// TIA Portal V19 export
FUNCTION "PID_DATA_MAPPING" : Void   // FC3, LAD
{ S7_Optimized_Access := 'TRUE' }
// stored: SetENOAutomatically false
BEGIN

REGION Network 1: -------------------------------------------------- REACTOR-1 ------------------------------------------------------------------
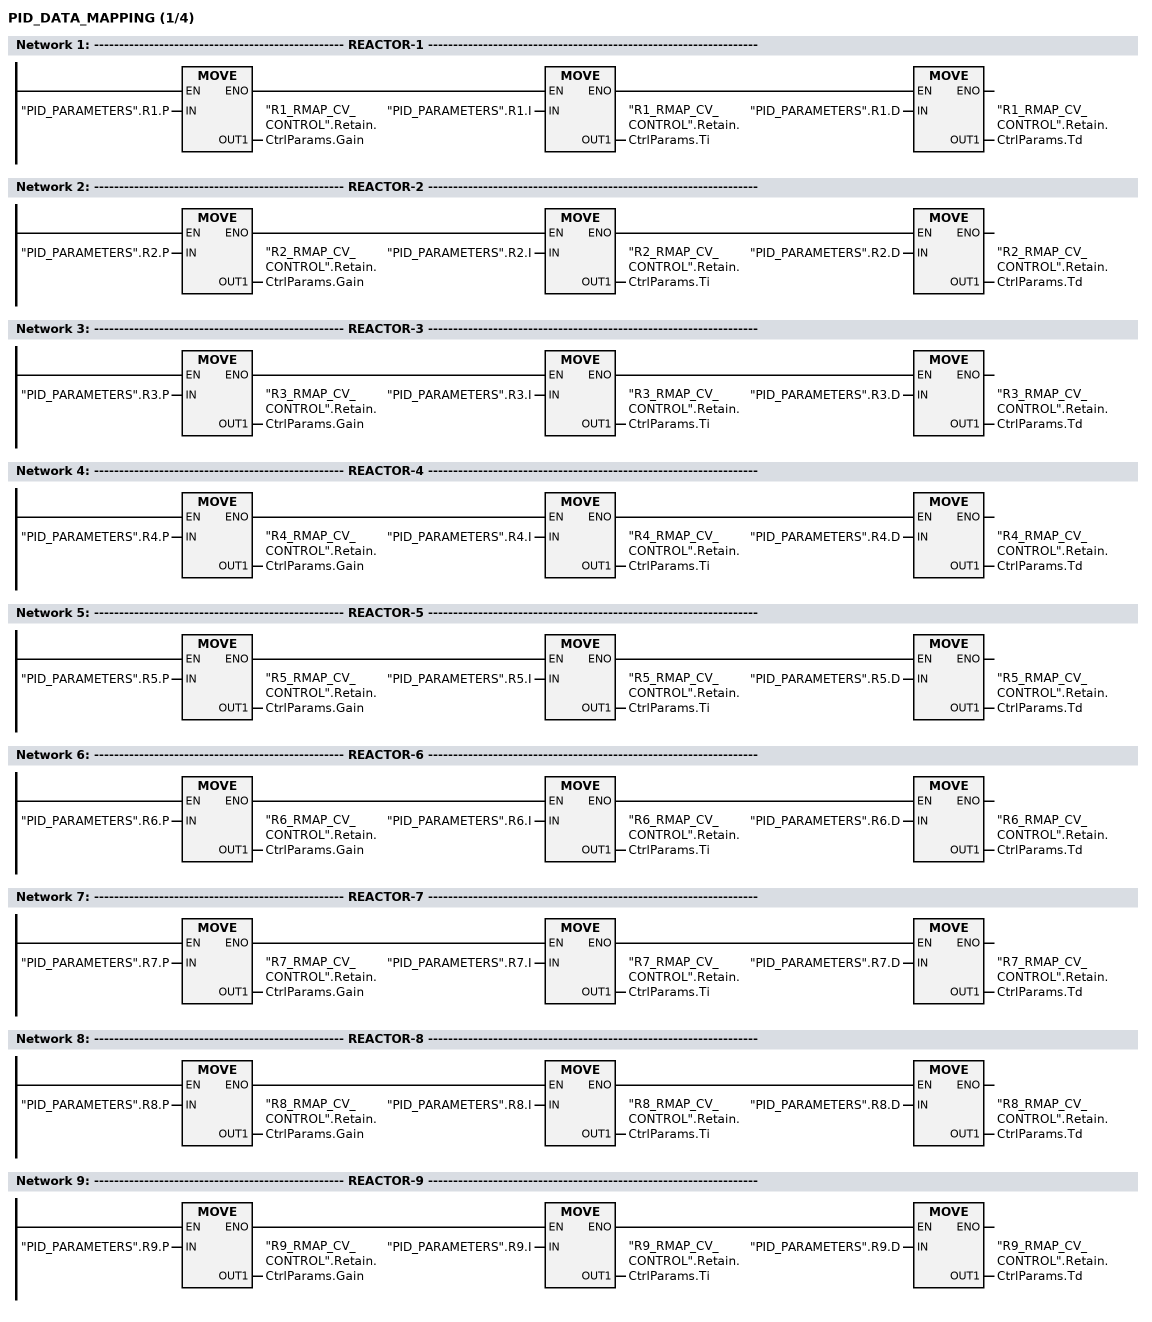
   RUNG wire#powerrail
      Move(in := "PID_PARAMETERS".R1.P, out1 => "R1_RMAP_CV_CONTROL".Retain.CtrlParams.Gain)
      Move(in := "PID_PARAMETERS".R1.I, out1 => "R1_RMAP_CV_CONTROL".Retain.CtrlParams.Ti)
      Move(in := "PID_PARAMETERS".R1.D, out1 => "R1_RMAP_CV_CONTROL".Retain.CtrlParams.Td)
   END_RUNG
   // the same network as SCL:
   "R1_RMAP_CV_CONTROL".Retain.CtrlParams.Gain := "PID_PARAMETERS".R1.P;
   "R1_RMAP_CV_CONTROL".Retain.CtrlParams.Ti := "PID_PARAMETERS".R1.I;
   "R1_RMAP_CV_CONTROL".Retain.CtrlParams.Td := "PID_PARAMETERS".R1.D;
END_REGION

REGION Network 2: -------------------------------------------------- REACTOR-2 ------------------------------------------------------------------
   RUNG wire#powerrail
      Move(in := "PID_PARAMETERS".R2.P, out1 => "R2_RMAP_CV_CONTROL".Retain.CtrlParams.Gain)
      Move(in := "PID_PARAMETERS".R2.I, out1 => "R2_RMAP_CV_CONTROL".Retain.CtrlParams.Ti)
      Move(in := "PID_PARAMETERS".R2.D, out1 => "R2_RMAP_CV_CONTROL".Retain.CtrlParams.Td)
   END_RUNG
   // the same network as SCL:
   "R2_RMAP_CV_CONTROL".Retain.CtrlParams.Gain := "PID_PARAMETERS".R2.P;
   "R2_RMAP_CV_CONTROL".Retain.CtrlParams.Ti := "PID_PARAMETERS".R2.I;
   "R2_RMAP_CV_CONTROL".Retain.CtrlParams.Td := "PID_PARAMETERS".R2.D;
END_REGION

REGION Network 3: -------------------------------------------------- REACTOR-3 ------------------------------------------------------------------
   RUNG wire#powerrail
      Move(in := "PID_PARAMETERS".R3.P, out1 => "R3_RMAP_CV_CONTROL".Retain.CtrlParams.Gain)
      Move(in := "PID_PARAMETERS".R3.I, out1 => "R3_RMAP_CV_CONTROL".Retain.CtrlParams.Ti)
      Move(in := "PID_PARAMETERS".R3.D, out1 => "R3_RMAP_CV_CONTROL".Retain.CtrlParams.Td)
   END_RUNG
   // the same network as SCL:
   "R3_RMAP_CV_CONTROL".Retain.CtrlParams.Gain := "PID_PARAMETERS".R3.P;
   "R3_RMAP_CV_CONTROL".Retain.CtrlParams.Ti := "PID_PARAMETERS".R3.I;
   "R3_RMAP_CV_CONTROL".Retain.CtrlParams.Td := "PID_PARAMETERS".R3.D;
END_REGION

REGION Network 4: -------------------------------------------------- REACTOR-4 ------------------------------------------------------------------
   RUNG wire#powerrail
      Move(in := "PID_PARAMETERS".R4.P, out1 => "R4_RMAP_CV_CONTROL".Retain.CtrlParams.Gain)
      Move(in := "PID_PARAMETERS".R4.I, out1 => "R4_RMAP_CV_CONTROL".Retain.CtrlParams.Ti)
      Move(in := "PID_PARAMETERS".R4.D, out1 => "R4_RMAP_CV_CONTROL".Retain.CtrlParams.Td)
   END_RUNG
   // the same network as SCL:
   "R4_RMAP_CV_CONTROL".Retain.CtrlParams.Gain := "PID_PARAMETERS".R4.P;
   "R4_RMAP_CV_CONTROL".Retain.CtrlParams.Ti := "PID_PARAMETERS".R4.I;
   "R4_RMAP_CV_CONTROL".Retain.CtrlParams.Td := "PID_PARAMETERS".R4.D;
END_REGION

REGION Network 5: -------------------------------------------------- REACTOR-5 ------------------------------------------------------------------
   RUNG wire#powerrail
      Move(in := "PID_PARAMETERS".R5.P, out1 => "R5_RMAP_CV_CONTROL".Retain.CtrlParams.Gain)
      Move(in := "PID_PARAMETERS".R5.I, out1 => "R5_RMAP_CV_CONTROL".Retain.CtrlParams.Ti)
      Move(in := "PID_PARAMETERS".R5.D, out1 => "R5_RMAP_CV_CONTROL".Retain.CtrlParams.Td)
   END_RUNG
   // the same network as SCL:
   "R5_RMAP_CV_CONTROL".Retain.CtrlParams.Gain := "PID_PARAMETERS".R5.P;
   "R5_RMAP_CV_CONTROL".Retain.CtrlParams.Ti := "PID_PARAMETERS".R5.I;
   "R5_RMAP_CV_CONTROL".Retain.CtrlParams.Td := "PID_PARAMETERS".R5.D;
END_REGION

REGION Network 6: -------------------------------------------------- REACTOR-6 ------------------------------------------------------------------
   RUNG wire#powerrail
      Move(in := "PID_PARAMETERS".R6.P, out1 => "R6_RMAP_CV_CONTROL".Retain.CtrlParams.Gain)
      Move(in := "PID_PARAMETERS".R6.I, out1 => "R6_RMAP_CV_CONTROL".Retain.CtrlParams.Ti)
      Move(in := "PID_PARAMETERS".R6.D, out1 => "R6_RMAP_CV_CONTROL".Retain.CtrlParams.Td)
   END_RUNG
   // the same network as SCL:
   "R6_RMAP_CV_CONTROL".Retain.CtrlParams.Gain := "PID_PARAMETERS".R6.P;
   "R6_RMAP_CV_CONTROL".Retain.CtrlParams.Ti := "PID_PARAMETERS".R6.I;
   "R6_RMAP_CV_CONTROL".Retain.CtrlParams.Td := "PID_PARAMETERS".R6.D;
END_REGION

REGION Network 7: -------------------------------------------------- REACTOR-7 ------------------------------------------------------------------
   RUNG wire#powerrail
      Move(in := "PID_PARAMETERS".R7.P, out1 => "R7_RMAP_CV_CONTROL".Retain.CtrlParams.Gain)
      Move(in := "PID_PARAMETERS".R7.I, out1 => "R7_RMAP_CV_CONTROL".Retain.CtrlParams.Ti)
      Move(in := "PID_PARAMETERS".R7.D, out1 => "R7_RMAP_CV_CONTROL".Retain.CtrlParams.Td)
   END_RUNG
   // the same network as SCL:
   "R7_RMAP_CV_CONTROL".Retain.CtrlParams.Gain := "PID_PARAMETERS".R7.P;
   "R7_RMAP_CV_CONTROL".Retain.CtrlParams.Ti := "PID_PARAMETERS".R7.I;
   "R7_RMAP_CV_CONTROL".Retain.CtrlParams.Td := "PID_PARAMETERS".R7.D;
END_REGION

REGION Network 8: -------------------------------------------------- REACTOR-8 ------------------------------------------------------------------
   RUNG wire#powerrail
      Move(in := "PID_PARAMETERS".R8.P, out1 => "R8_RMAP_CV_CONTROL".Retain.CtrlParams.Gain)
      Move(in := "PID_PARAMETERS".R8.I, out1 => "R8_RMAP_CV_CONTROL".Retain.CtrlParams.Ti)
      Move(in := "PID_PARAMETERS".R8.D, out1 => "R8_RMAP_CV_CONTROL".Retain.CtrlParams.Td)
   END_RUNG
   // the same network as SCL:
   "R8_RMAP_CV_CONTROL".Retain.CtrlParams.Gain := "PID_PARAMETERS".R8.P;
   "R8_RMAP_CV_CONTROL".Retain.CtrlParams.Ti := "PID_PARAMETERS".R8.I;
   "R8_RMAP_CV_CONTROL".Retain.CtrlParams.Td := "PID_PARAMETERS".R8.D;
END_REGION

REGION Network 9: -------------------------------------------------- REACTOR-9 ------------------------------------------------------------------
   RUNG wire#powerrail
      Move(in := "PID_PARAMETERS".R9.P, out1 => "R9_RMAP_CV_CONTROL".Retain.CtrlParams.Gain)
      Move(in := "PID_PARAMETERS".R9.I, out1 => "R9_RMAP_CV_CONTROL".Retain.CtrlParams.Ti)
      Move(in := "PID_PARAMETERS".R9.D, out1 => "R9_RMAP_CV_CONTROL".Retain.CtrlParams.Td)
   END_RUNG
   // the same network as SCL:
   "R9_RMAP_CV_CONTROL".Retain.CtrlParams.Gain := "PID_PARAMETERS".R9.P;
   "R9_RMAP_CV_CONTROL".Retain.CtrlParams.Ti := "PID_PARAMETERS".R9.I;
   "R9_RMAP_CV_CONTROL".Retain.CtrlParams.Td := "PID_PARAMETERS".R9.D;
END_REGION

REGION Network 10: -------------------------------------------------- REACTOR-10 ------------------------------------------------------------------
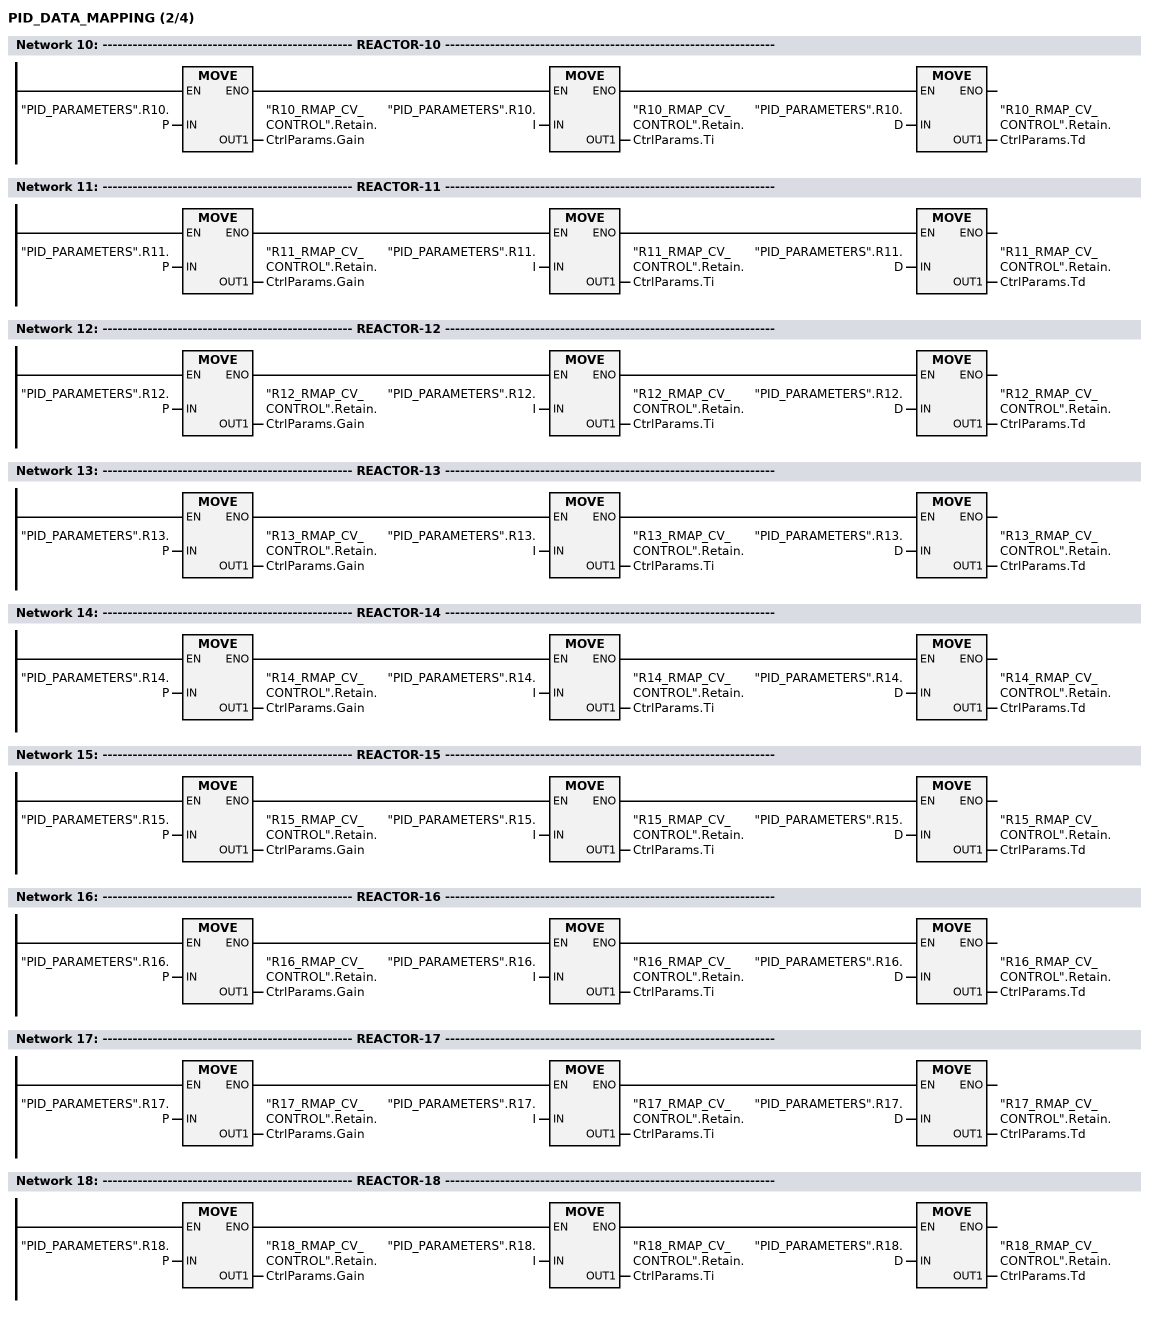
   RUNG wire#powerrail
      Move(in := "PID_PARAMETERS".R10.P, out1 => "R10_RMAP_CV_CONTROL".Retain.CtrlParams.Gain)
      Move(in := "PID_PARAMETERS".R10.I, out1 => "R10_RMAP_CV_CONTROL".Retain.CtrlParams.Ti)
      Move(in := "PID_PARAMETERS".R10.D, out1 => "R10_RMAP_CV_CONTROL".Retain.CtrlParams.Td)
   END_RUNG
   // the same network as SCL:
   "R10_RMAP_CV_CONTROL".Retain.CtrlParams.Gain := "PID_PARAMETERS".R10.P;
   "R10_RMAP_CV_CONTROL".Retain.CtrlParams.Ti := "PID_PARAMETERS".R10.I;
   "R10_RMAP_CV_CONTROL".Retain.CtrlParams.Td := "PID_PARAMETERS".R10.D;
END_REGION

REGION Network 11: -------------------------------------------------- REACTOR-11 ------------------------------------------------------------------
   RUNG wire#powerrail
      Move(in := "PID_PARAMETERS".R11.P, out1 => "R11_RMAP_CV_CONTROL".Retain.CtrlParams.Gain)
      Move(in := "PID_PARAMETERS".R11.I, out1 => "R11_RMAP_CV_CONTROL".Retain.CtrlParams.Ti)
      Move(in := "PID_PARAMETERS".R11.D, out1 => "R11_RMAP_CV_CONTROL".Retain.CtrlParams.Td)
   END_RUNG
   // the same network as SCL:
   "R11_RMAP_CV_CONTROL".Retain.CtrlParams.Gain := "PID_PARAMETERS".R11.P;
   "R11_RMAP_CV_CONTROL".Retain.CtrlParams.Ti := "PID_PARAMETERS".R11.I;
   "R11_RMAP_CV_CONTROL".Retain.CtrlParams.Td := "PID_PARAMETERS".R11.D;
END_REGION

REGION Network 12: -------------------------------------------------- REACTOR-12 ------------------------------------------------------------------
   RUNG wire#powerrail
      Move(in := "PID_PARAMETERS".R12.P, out1 => "R12_RMAP_CV_CONTROL".Retain.CtrlParams.Gain)
      Move(in := "PID_PARAMETERS".R12.I, out1 => "R12_RMAP_CV_CONTROL".Retain.CtrlParams.Ti)
      Move(in := "PID_PARAMETERS".R12.D, out1 => "R12_RMAP_CV_CONTROL".Retain.CtrlParams.Td)
   END_RUNG
   // the same network as SCL:
   "R12_RMAP_CV_CONTROL".Retain.CtrlParams.Gain := "PID_PARAMETERS".R12.P;
   "R12_RMAP_CV_CONTROL".Retain.CtrlParams.Ti := "PID_PARAMETERS".R12.I;
   "R12_RMAP_CV_CONTROL".Retain.CtrlParams.Td := "PID_PARAMETERS".R12.D;
END_REGION

REGION Network 13: -------------------------------------------------- REACTOR-13 ------------------------------------------------------------------
   RUNG wire#powerrail
      Move(in := "PID_PARAMETERS".R13.P, out1 => "R13_RMAP_CV_CONTROL".Retain.CtrlParams.Gain)
      Move(in := "PID_PARAMETERS".R13.I, out1 => "R13_RMAP_CV_CONTROL".Retain.CtrlParams.Ti)
      Move(in := "PID_PARAMETERS".R13.D, out1 => "R13_RMAP_CV_CONTROL".Retain.CtrlParams.Td)
   END_RUNG
   // the same network as SCL:
   "R13_RMAP_CV_CONTROL".Retain.CtrlParams.Gain := "PID_PARAMETERS".R13.P;
   "R13_RMAP_CV_CONTROL".Retain.CtrlParams.Ti := "PID_PARAMETERS".R13.I;
   "R13_RMAP_CV_CONTROL".Retain.CtrlParams.Td := "PID_PARAMETERS".R13.D;
END_REGION

REGION Network 14: -------------------------------------------------- REACTOR-14 ------------------------------------------------------------------
   RUNG wire#powerrail
      Move(in := "PID_PARAMETERS".R14.P, out1 => "R14_RMAP_CV_CONTROL".Retain.CtrlParams.Gain)
      Move(in := "PID_PARAMETERS".R14.I, out1 => "R14_RMAP_CV_CONTROL".Retain.CtrlParams.Ti)
      Move(in := "PID_PARAMETERS".R14.D, out1 => "R14_RMAP_CV_CONTROL".Retain.CtrlParams.Td)
   END_RUNG
   // the same network as SCL:
   "R14_RMAP_CV_CONTROL".Retain.CtrlParams.Gain := "PID_PARAMETERS".R14.P;
   "R14_RMAP_CV_CONTROL".Retain.CtrlParams.Ti := "PID_PARAMETERS".R14.I;
   "R14_RMAP_CV_CONTROL".Retain.CtrlParams.Td := "PID_PARAMETERS".R14.D;
END_REGION

REGION Network 15: -------------------------------------------------- REACTOR-15 ------------------------------------------------------------------
   RUNG wire#powerrail
      Move(in := "PID_PARAMETERS".R15.P, out1 => "R15_RMAP_CV_CONTROL".Retain.CtrlParams.Gain)
      Move(in := "PID_PARAMETERS".R15.I, out1 => "R15_RMAP_CV_CONTROL".Retain.CtrlParams.Ti)
      Move(in := "PID_PARAMETERS".R15.D, out1 => "R15_RMAP_CV_CONTROL".Retain.CtrlParams.Td)
   END_RUNG
   // the same network as SCL:
   "R15_RMAP_CV_CONTROL".Retain.CtrlParams.Gain := "PID_PARAMETERS".R15.P;
   "R15_RMAP_CV_CONTROL".Retain.CtrlParams.Ti := "PID_PARAMETERS".R15.I;
   "R15_RMAP_CV_CONTROL".Retain.CtrlParams.Td := "PID_PARAMETERS".R15.D;
END_REGION

REGION Network 16: -------------------------------------------------- REACTOR-16 ------------------------------------------------------------------
   RUNG wire#powerrail
      Move(in := "PID_PARAMETERS".R16.P, out1 => "R16_RMAP_CV_CONTROL".Retain.CtrlParams.Gain)
      Move(in := "PID_PARAMETERS".R16.I, out1 => "R16_RMAP_CV_CONTROL".Retain.CtrlParams.Ti)
      Move(in := "PID_PARAMETERS".R16.D, out1 => "R16_RMAP_CV_CONTROL".Retain.CtrlParams.Td)
   END_RUNG
   // the same network as SCL:
   "R16_RMAP_CV_CONTROL".Retain.CtrlParams.Gain := "PID_PARAMETERS".R16.P;
   "R16_RMAP_CV_CONTROL".Retain.CtrlParams.Ti := "PID_PARAMETERS".R16.I;
   "R16_RMAP_CV_CONTROL".Retain.CtrlParams.Td := "PID_PARAMETERS".R16.D;
END_REGION

REGION Network 17: -------------------------------------------------- REACTOR-17 ------------------------------------------------------------------
   RUNG wire#powerrail
      Move(in := "PID_PARAMETERS".R17.P, out1 => "R17_RMAP_CV_CONTROL".Retain.CtrlParams.Gain)
      Move(in := "PID_PARAMETERS".R17.I, out1 => "R17_RMAP_CV_CONTROL".Retain.CtrlParams.Ti)
      Move(in := "PID_PARAMETERS".R17.D, out1 => "R17_RMAP_CV_CONTROL".Retain.CtrlParams.Td)
   END_RUNG
   // the same network as SCL:
   "R17_RMAP_CV_CONTROL".Retain.CtrlParams.Gain := "PID_PARAMETERS".R17.P;
   "R17_RMAP_CV_CONTROL".Retain.CtrlParams.Ti := "PID_PARAMETERS".R17.I;
   "R17_RMAP_CV_CONTROL".Retain.CtrlParams.Td := "PID_PARAMETERS".R17.D;
END_REGION

REGION Network 18: -------------------------------------------------- REACTOR-18 ------------------------------------------------------------------
   RUNG wire#powerrail
      Move(in := "PID_PARAMETERS".R18.P, out1 => "R18_RMAP_CV_CONTROL".Retain.CtrlParams.Gain)
      Move(in := "PID_PARAMETERS".R18.I, out1 => "R18_RMAP_CV_CONTROL".Retain.CtrlParams.Ti)
      Move(in := "PID_PARAMETERS".R18.D, out1 => "R18_RMAP_CV_CONTROL".Retain.CtrlParams.Td)
   END_RUNG
   // the same network as SCL:
   "R18_RMAP_CV_CONTROL".Retain.CtrlParams.Gain := "PID_PARAMETERS".R18.P;
   "R18_RMAP_CV_CONTROL".Retain.CtrlParams.Ti := "PID_PARAMETERS".R18.I;
   "R18_RMAP_CV_CONTROL".Retain.CtrlParams.Td := "PID_PARAMETERS".R18.D;
END_REGION

REGION Network 19: -------------------------------------------------- HS_CP01 ------------------------------------------------------------------
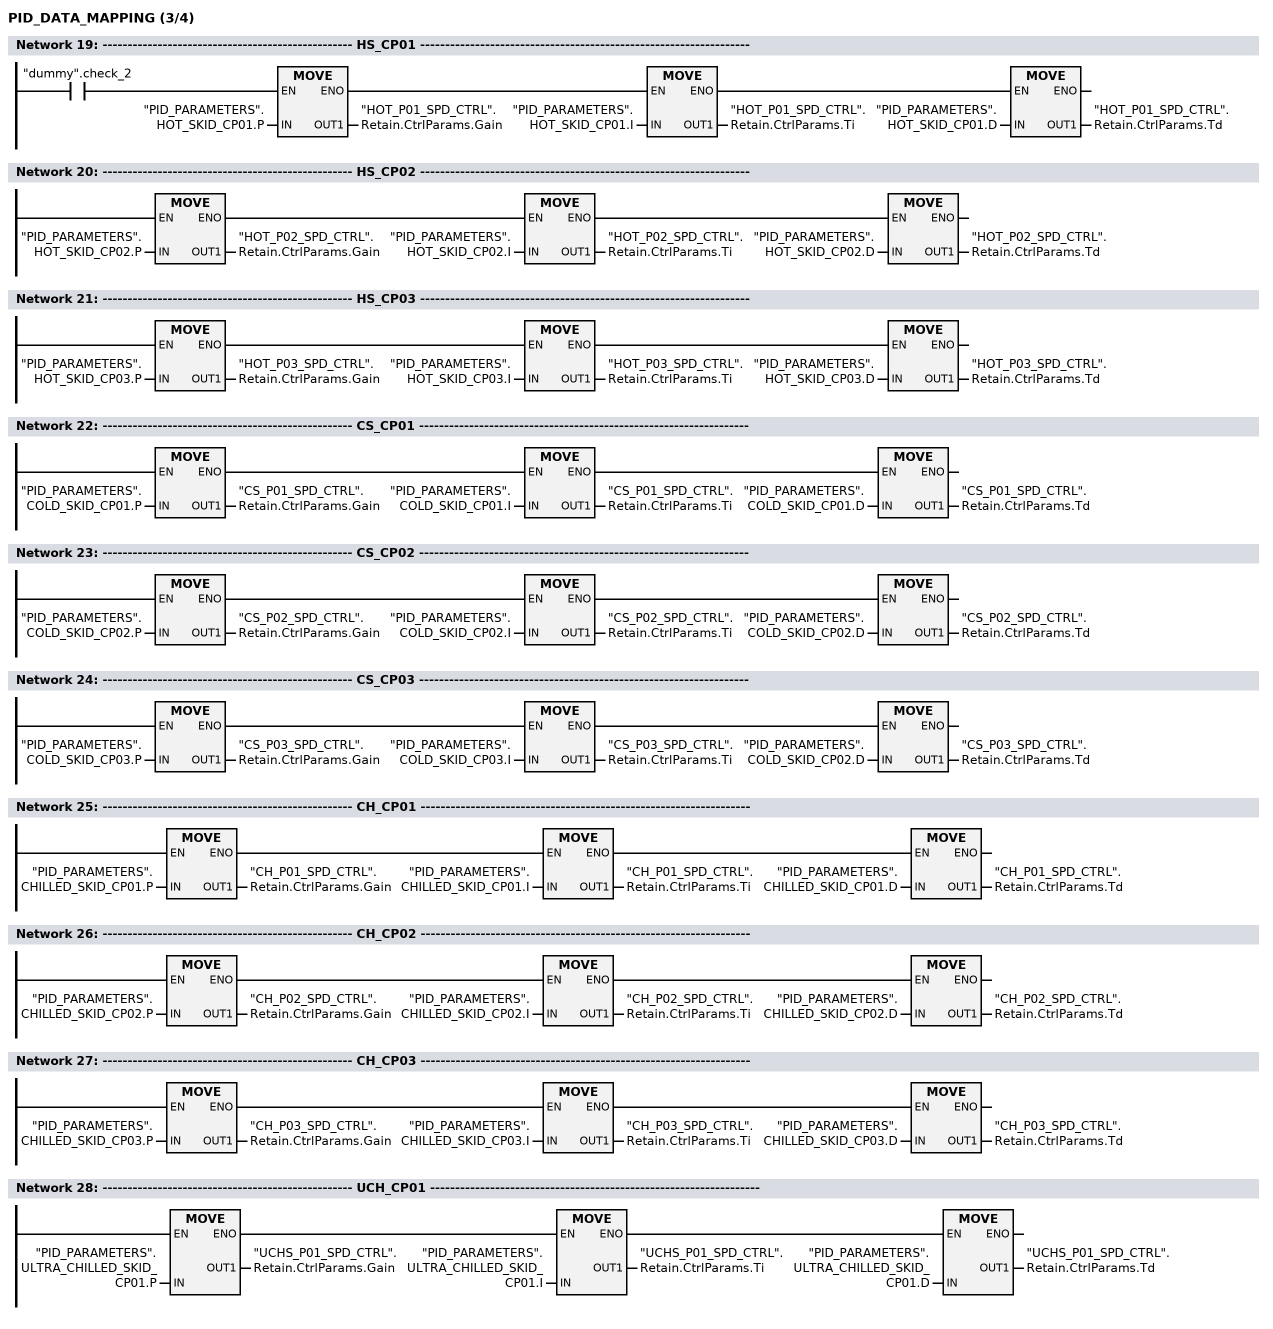
   RUNG wire#powerrail
      Contact( "dummy".check_2 )
      Move(in := "PID_PARAMETERS".HOT_SKID_CP01.P, out1 => "HOT_P01_SPD_CTRL".Retain.CtrlParams.Gain)
      Move(in := "PID_PARAMETERS".HOT_SKID_CP01.I, out1 => "HOT_P01_SPD_CTRL".Retain.CtrlParams.Ti)
      Move(in := "PID_PARAMETERS".HOT_SKID_CP01.D, out1 => "HOT_P01_SPD_CTRL".Retain.CtrlParams.Td)
   END_RUNG
   // the same network as SCL:
   IF "dummy".check_2 THEN
       "HOT_P01_SPD_CTRL".Retain.CtrlParams.Gain := "PID_PARAMETERS".HOT_SKID_CP01.P;
       "HOT_P01_SPD_CTRL".Retain.CtrlParams.Ti := "PID_PARAMETERS".HOT_SKID_CP01.I;
       "HOT_P01_SPD_CTRL".Retain.CtrlParams.Td := "PID_PARAMETERS".HOT_SKID_CP01.D;
   END_IF;
END_REGION

REGION Network 20: -------------------------------------------------- HS_CP02 ------------------------------------------------------------------
   RUNG wire#powerrail
      Move(in := "PID_PARAMETERS".HOT_SKID_CP02.P, out1 => "HOT_P02_SPD_CTRL".Retain.CtrlParams.Gain)
      Move(in := "PID_PARAMETERS".HOT_SKID_CP02.I, out1 => "HOT_P02_SPD_CTRL".Retain.CtrlParams.Ti)
      Move(in := "PID_PARAMETERS".HOT_SKID_CP02.D, out1 => "HOT_P02_SPD_CTRL".Retain.CtrlParams.Td)
   END_RUNG
   // the same network as SCL:
   "HOT_P02_SPD_CTRL".Retain.CtrlParams.Gain := "PID_PARAMETERS".HOT_SKID_CP02.P;
   "HOT_P02_SPD_CTRL".Retain.CtrlParams.Ti := "PID_PARAMETERS".HOT_SKID_CP02.I;
   "HOT_P02_SPD_CTRL".Retain.CtrlParams.Td := "PID_PARAMETERS".HOT_SKID_CP02.D;
END_REGION

REGION Network 21: -------------------------------------------------- HS_CP03 ------------------------------------------------------------------
   RUNG wire#powerrail
      Move(in := "PID_PARAMETERS".HOT_SKID_CP03.P, out1 => "HOT_P03_SPD_CTRL".Retain.CtrlParams.Gain)
      Move(in := "PID_PARAMETERS".HOT_SKID_CP03.I, out1 => "HOT_P03_SPD_CTRL".Retain.CtrlParams.Ti)
      Move(in := "PID_PARAMETERS".HOT_SKID_CP03.D, out1 => "HOT_P03_SPD_CTRL".Retain.CtrlParams.Td)
   END_RUNG
   // the same network as SCL:
   "HOT_P03_SPD_CTRL".Retain.CtrlParams.Gain := "PID_PARAMETERS".HOT_SKID_CP03.P;
   "HOT_P03_SPD_CTRL".Retain.CtrlParams.Ti := "PID_PARAMETERS".HOT_SKID_CP03.I;
   "HOT_P03_SPD_CTRL".Retain.CtrlParams.Td := "PID_PARAMETERS".HOT_SKID_CP03.D;
END_REGION

REGION Network 22: -------------------------------------------------- CS_CP01 ------------------------------------------------------------------
   RUNG wire#powerrail
      Move(in := "PID_PARAMETERS".COLD_SKID_CP01.P, out1 => "CS_P01_SPD_CTRL".Retain.CtrlParams.Gain)
      Move(in := "PID_PARAMETERS".COLD_SKID_CP01.I, out1 => "CS_P01_SPD_CTRL".Retain.CtrlParams.Ti)
      Move(in := "PID_PARAMETERS".COLD_SKID_CP01.D, out1 => "CS_P01_SPD_CTRL".Retain.CtrlParams.Td)
   END_RUNG
   // the same network as SCL:
   "CS_P01_SPD_CTRL".Retain.CtrlParams.Gain := "PID_PARAMETERS".COLD_SKID_CP01.P;
   "CS_P01_SPD_CTRL".Retain.CtrlParams.Ti := "PID_PARAMETERS".COLD_SKID_CP01.I;
   "CS_P01_SPD_CTRL".Retain.CtrlParams.Td := "PID_PARAMETERS".COLD_SKID_CP01.D;
END_REGION

REGION Network 23: -------------------------------------------------- CS_CP02 ------------------------------------------------------------------
   RUNG wire#powerrail
      Move(in := "PID_PARAMETERS".COLD_SKID_CP02.P, out1 => "CS_P02_SPD_CTRL".Retain.CtrlParams.Gain)
      Move(in := "PID_PARAMETERS".COLD_SKID_CP02.I, out1 => "CS_P02_SPD_CTRL".Retain.CtrlParams.Ti)
      Move(in := "PID_PARAMETERS".COLD_SKID_CP02.D, out1 => "CS_P02_SPD_CTRL".Retain.CtrlParams.Td)
   END_RUNG
   // the same network as SCL:
   "CS_P02_SPD_CTRL".Retain.CtrlParams.Gain := "PID_PARAMETERS".COLD_SKID_CP02.P;
   "CS_P02_SPD_CTRL".Retain.CtrlParams.Ti := "PID_PARAMETERS".COLD_SKID_CP02.I;
   "CS_P02_SPD_CTRL".Retain.CtrlParams.Td := "PID_PARAMETERS".COLD_SKID_CP02.D;
END_REGION

REGION Network 24: -------------------------------------------------- CS_CP03 ------------------------------------------------------------------
   RUNG wire#powerrail
      Move(in := "PID_PARAMETERS".COLD_SKID_CP03.P, out1 => "CS_P03_SPD_CTRL".Retain.CtrlParams.Gain)
      Move(in := "PID_PARAMETERS".COLD_SKID_CP03.I, out1 => "CS_P03_SPD_CTRL".Retain.CtrlParams.Ti)
      Move(in := "PID_PARAMETERS".COLD_SKID_CP02.D, out1 => "CS_P03_SPD_CTRL".Retain.CtrlParams.Td)
   END_RUNG
   // the same network as SCL:
   "CS_P03_SPD_CTRL".Retain.CtrlParams.Gain := "PID_PARAMETERS".COLD_SKID_CP03.P;
   "CS_P03_SPD_CTRL".Retain.CtrlParams.Ti := "PID_PARAMETERS".COLD_SKID_CP03.I;
   "CS_P03_SPD_CTRL".Retain.CtrlParams.Td := "PID_PARAMETERS".COLD_SKID_CP02.D;
END_REGION

REGION Network 25: -------------------------------------------------- CH_CP01 ------------------------------------------------------------------
   RUNG wire#powerrail
      Move(in := "PID_PARAMETERS".CHILLED_SKID_CP01.P, out1 => "CH_P01_SPD_CTRL".Retain.CtrlParams.Gain)
      Move(in := "PID_PARAMETERS".CHILLED_SKID_CP01.I, out1 => "CH_P01_SPD_CTRL".Retain.CtrlParams.Ti)
      Move(in := "PID_PARAMETERS".CHILLED_SKID_CP01.D, out1 => "CH_P01_SPD_CTRL".Retain.CtrlParams.Td)
   END_RUNG
   // the same network as SCL:
   "CH_P01_SPD_CTRL".Retain.CtrlParams.Gain := "PID_PARAMETERS".CHILLED_SKID_CP01.P;
   "CH_P01_SPD_CTRL".Retain.CtrlParams.Ti := "PID_PARAMETERS".CHILLED_SKID_CP01.I;
   "CH_P01_SPD_CTRL".Retain.CtrlParams.Td := "PID_PARAMETERS".CHILLED_SKID_CP01.D;
END_REGION

REGION Network 26: -------------------------------------------------- CH_CP02 ------------------------------------------------------------------
   RUNG wire#powerrail
      Move(in := "PID_PARAMETERS".CHILLED_SKID_CP02.P, out1 => "CH_P02_SPD_CTRL".Retain.CtrlParams.Gain)
      Move(in := "PID_PARAMETERS".CHILLED_SKID_CP02.I, out1 => "CH_P02_SPD_CTRL".Retain.CtrlParams.Ti)
      Move(in := "PID_PARAMETERS".CHILLED_SKID_CP02.D, out1 => "CH_P02_SPD_CTRL".Retain.CtrlParams.Td)
   END_RUNG
   // the same network as SCL:
   "CH_P02_SPD_CTRL".Retain.CtrlParams.Gain := "PID_PARAMETERS".CHILLED_SKID_CP02.P;
   "CH_P02_SPD_CTRL".Retain.CtrlParams.Ti := "PID_PARAMETERS".CHILLED_SKID_CP02.I;
   "CH_P02_SPD_CTRL".Retain.CtrlParams.Td := "PID_PARAMETERS".CHILLED_SKID_CP02.D;
END_REGION

REGION Network 27: -------------------------------------------------- CH_CP03 ------------------------------------------------------------------
   RUNG wire#powerrail
      Move(in := "PID_PARAMETERS".CHILLED_SKID_CP03.P, out1 => "CH_P03_SPD_CTRL".Retain.CtrlParams.Gain)
      Move(in := "PID_PARAMETERS".CHILLED_SKID_CP03.I, out1 => "CH_P03_SPD_CTRL".Retain.CtrlParams.Ti)
      Move(in := "PID_PARAMETERS".CHILLED_SKID_CP03.D, out1 => "CH_P03_SPD_CTRL".Retain.CtrlParams.Td)
   END_RUNG
   // the same network as SCL:
   "CH_P03_SPD_CTRL".Retain.CtrlParams.Gain := "PID_PARAMETERS".CHILLED_SKID_CP03.P;
   "CH_P03_SPD_CTRL".Retain.CtrlParams.Ti := "PID_PARAMETERS".CHILLED_SKID_CP03.I;
   "CH_P03_SPD_CTRL".Retain.CtrlParams.Td := "PID_PARAMETERS".CHILLED_SKID_CP03.D;
END_REGION

REGION Network 28: -------------------------------------------------- UCH_CP01 ------------------------------------------------------------------
   RUNG wire#powerrail
      Move(in := "PID_PARAMETERS".ULTRA_CHILLED_SKID_CP01.P, out1 => "UCHS_P01_SPD_CTRL".Retain.CtrlParams.Gain)
      Move(in := "PID_PARAMETERS".ULTRA_CHILLED_SKID_CP01.I, out1 => "UCHS_P01_SPD_CTRL".Retain.CtrlParams.Ti)
      Move(in := "PID_PARAMETERS".ULTRA_CHILLED_SKID_CP01.D, out1 => "UCHS_P01_SPD_CTRL".Retain.CtrlParams.Td)
   END_RUNG
   // the same network as SCL:
   "UCHS_P01_SPD_CTRL".Retain.CtrlParams.Gain := "PID_PARAMETERS".ULTRA_CHILLED_SKID_CP01.P;
   "UCHS_P01_SPD_CTRL".Retain.CtrlParams.Ti := "PID_PARAMETERS".ULTRA_CHILLED_SKID_CP01.I;
   "UCHS_P01_SPD_CTRL".Retain.CtrlParams.Td := "PID_PARAMETERS".ULTRA_CHILLED_SKID_CP01.D;
END_REGION

REGION Network 29: -------------------------------------------------- UCH_CP02 ------------------------------------------------------------------
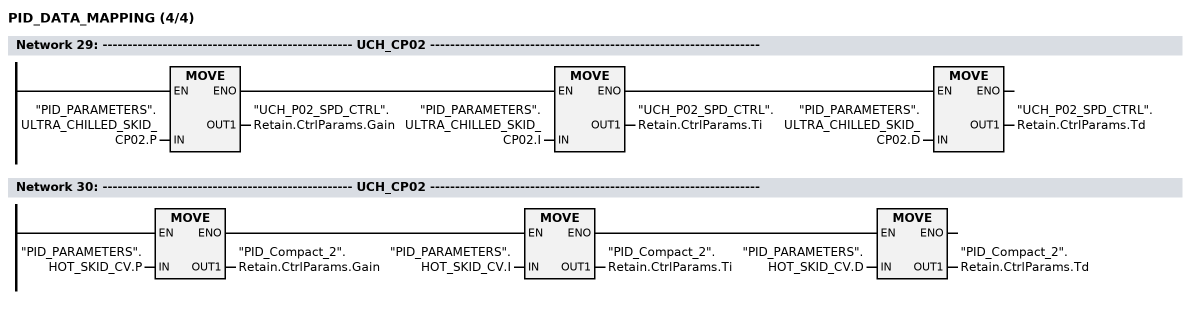
   RUNG wire#powerrail
      Move(in := "PID_PARAMETERS".ULTRA_CHILLED_SKID_CP02.P, out1 => "UCH_P02_SPD_CTRL".Retain.CtrlParams.Gain)
      Move(in := "PID_PARAMETERS".ULTRA_CHILLED_SKID_CP02.I, out1 => "UCH_P02_SPD_CTRL".Retain.CtrlParams.Ti)
      Move(in := "PID_PARAMETERS".ULTRA_CHILLED_SKID_CP02.D, out1 => "UCH_P02_SPD_CTRL".Retain.CtrlParams.Td)
   END_RUNG
   // the same network as SCL:
   "UCH_P02_SPD_CTRL".Retain.CtrlParams.Gain := "PID_PARAMETERS".ULTRA_CHILLED_SKID_CP02.P;
   "UCH_P02_SPD_CTRL".Retain.CtrlParams.Ti := "PID_PARAMETERS".ULTRA_CHILLED_SKID_CP02.I;
   "UCH_P02_SPD_CTRL".Retain.CtrlParams.Td := "PID_PARAMETERS".ULTRA_CHILLED_SKID_CP02.D;
END_REGION

REGION Network 30: -------------------------------------------------- UCH_CP02 ------------------------------------------------------------------
   RUNG wire#powerrail
      Move(in := "PID_PARAMETERS".HOT_SKID_CV.P, out1 => "PID_Compact_2".Retain.CtrlParams.Gain)
      Move(in := "PID_PARAMETERS".HOT_SKID_CV.I, out1 => "PID_Compact_2".Retain.CtrlParams.Ti)
      Move(in := "PID_PARAMETERS".HOT_SKID_CV.D, out1 => "PID_Compact_2".Retain.CtrlParams.Td)
   END_RUNG
   // the same network as SCL:
   "PID_Compact_2".Retain.CtrlParams.Gain := "PID_PARAMETERS".HOT_SKID_CV.P;
   "PID_Compact_2".Retain.CtrlParams.Ti := "PID_PARAMETERS".HOT_SKID_CV.I;
   "PID_Compact_2".Retain.CtrlParams.Td := "PID_PARAMETERS".HOT_SKID_CV.D;
END_REGION
END_FUNCTION
